Staubli VAL3: putMessage.pgx

public program putMessage(string x_sMsg, string x_sMsgType)
begin
  switch x_sMsgType
    case "info"
      utTxt_popUpMsg.Appearance.sBackgroundColour="#7C95FF"
    break
    //
    case "warning"
      utTxt_popUpMsg.Appearance.sBackgroundColour="#EEFB45"
    break
    //
    case "confirm"
      utTxt_popUpMsg.Appearance.sBackgroundColour="#FFFFFF"
    break
    //
    default
      utTxt_popUpMsg.Appearance.sBackgroundColour="#ADADB2"
    break
  endSwitch
  utTxt_popUpMsg.Common.sValue=x_sMsg
  delay(0.2)
  utCtn_Message.Appearance.bVisibility=true
end
